(* IEC 61131-3 sources: sis-interlock-demo/pytests/golden/mini/src/GVLs/Generated, 3 files *)

(* ---- GVL_Sis.gvl.st ---- *)
// AUTO-GENERATED by cemgen 1.0.0 — не редактировать: правьте матрицу и запустите
//   python -m cemgen generate <файл матрицы .csv или .xlsx>
// Матрица: TEST-U301-CEM, объект U-301, ревизия 1 от 2026-10-16, SHA-256 сетки 9067fda96ae55e67
// Назначение: экземпляры ПАЗ объекта U-301: источник времени, журнал событий, приложение ПАЗ и
//             команды HMI (ST_SisCmd). Вызов — PRG_Sis.
// Автор:      pytest; код — генератор cemgen
// Версия:     1.0.0
// Документ:   docs/DESIGN.md, раздел «10. Генератор cemgen»; docs/cause_effect_matrix.md
// ВНИМАНИЕ:   код демонстрационный и не предназначен для систем безопасности. Реальная ПАЗ требует
//             определения SIL, сертифицированных аппаратных и программных средств и валидации по
//             ГОСТ Р МЭК 61511.
{attribute 'qualified_only'}
VAR_GLOBAL
    fbTime : PL.FB_SystemTime;   // монотонное время LTIME (PL.I_TimeSource)
    fbLog  : FB_SisEventLog;     // журнал событий ПАЗ, кольцо GVL_Const.SIS_LOG_SIZE
    fbApp  : FB_SisApp;          // ПАЗ объекта: привязка, голосование, матрица, выходы
    stCmd  : ST_SisCmd;          // команды HMI: сброс, пусковые обходы, байпасы каналов
END_VAR

(* ---- GVL_SisCfg.gvl.st ---- *)
// AUTO-GENERATED by cemgen 1.0.0 — не редактировать: правьте матрицу и запустите
//   python -m cemgen generate <файл матрицы .csv или .xlsx>
// Матрица: TEST-U301-CEM, объект U-301, ревизия 1 от 2026-10-16, SHA-256 сетки 9067fda96ae55e67
// Назначение: конфигурация ПАЗ объекта U-301 из матрицы причин и следствий: номера причин и
//             следствий, шкалы датчиков, матрица CEM_CFG (с CRC) и группы голосования VOTE_CFG.
//             VAR_GLOBAL CONSTANT: с HMI не меняется (решение D-09), правка — только через матрицу
//             и генератор.
// Автор:      pytest; код — генератор cemgen
// Версия:     1.0.0
// Документ:   docs/DESIGN.md, раздел «10. Генератор cemgen»; docs/cause_effect_matrix.md
// ВНИМАНИЕ:   код демонстрационный и не предназначен для систем безопасности. Реальная ПАЗ требует
//             определения SIL, сертифицированных аппаратных и программных средств и валидации по
//             ГОСТ Р МЭК 61511.
{attribute 'qualified_only'}
VAR_GLOBAL CONSTANT
    // Номера причин: индекс i строки матрицы, бит маски i − 1
    CAUSE_TSH301       : UINT := 1;   // Температура высокая
    CAUSE_PSL302       : UINT := 2;   // Давление низкое
    CAUSE_XS303        : UINT := 3;   // Внешний останов
    CAUSE_COUNT        : UINT := 3;   // причин в матрице
    // Номера следствий: индекс j столбца матрицы
    EFFECT_XV301       : UINT := 1;   // Отсечной клапан XV301
    EFFECT_M302        : UINT := 2;   // Насос M302
    EFFECT_COUNT       : UINT := 2;   // следствий в матрице
    // Шкалы датчиков 4–20 мА (инж. ед.) и нормальные токи для демо и тестов
    AI_TT301_LO_EU     : REAL := 0.0;   // TT301: шкала 0…100 °C
    AI_TT301_HI_EU     : REAL := 100.0;
    AI_TT301_NORMAL_MA : REAL := 10.4;   // 40 °C
    // Матрица причин и следствий (DESIGN.md, 4.2, 6.8): маска следствия — «X» в его столбце
    CEM_CFG : ST_CemCfg := (uiCauseCount := 3, uiEffectCount := 2, xStartTripped := FALSE,
        wMatrixCrc := 16#0F15,
        astCause := [
            (xEnable := TRUE, eSource := E_CauseSource.Voting, tDelay := T#1S),                 // 1 TSH301
            (xEnable := TRUE, eSource := E_CauseSource.Voting, tDelay := T#0S,
                xOverrideAllowed := TRUE, tOverrideMax := T#10M, tOverrideClear := T#30S),      // 2 PSL302
            (xEnable := TRUE, eSource := E_CauseSource.External, tDelay := T#500MS),            // 3 XS303
            (xEnable := FALSE),                                                                 // 4 — резерв
            (xEnable := FALSE),                                                                 // 5 — резерв
            (xEnable := FALSE),                                                                 // 6 — резерв
            (xEnable := FALSE),                                                                 // 7 — резерв
            (xEnable := FALSE),                                                                 // 8 — резерв
            (xEnable := FALSE),                                                                 // 9 — резерв
            (xEnable := FALSE),                                                                 // 10 — резерв
            (xEnable := FALSE),                                                                 // 11 — резерв
            (xEnable := FALSE),                                                                 // 12 — резерв
            (xEnable := FALSE),                                                                 // 13 — резерв
            (xEnable := FALSE),                                                                 // 14 — резерв
            (xEnable := FALSE),                                                                 // 15 — резерв
            (xEnable := FALSE)],                                                                // 16 — резерв
        astEffect := [
            (eSafeState := E_SafeState.Closed, wCauseMask := 16#0003),                          // 1 XV301: 1, 2
            (eSafeState := E_SafeState.Stopped, wCauseMask := 16#0006),                         // 2 M302: 2, 3
            (wCauseMask := 0),                                                                  // 3 — резерв
            (wCauseMask := 0),                                                                  // 4 — резерв
            (wCauseMask := 0),                                                                  // 5 — резерв
            (wCauseMask := 0),                                                                  // 6 — резерв
            (wCauseMask := 0),                                                                  // 7 — резерв
            (wCauseMask := 0),                                                                  // 8 — резерв
            (wCauseMask := 0),                                                                  // 9 — резерв
            (wCauseMask := 0),                                                                  // 10 — резерв
            (wCauseMask := 0),                                                                  // 11 — резерв
            (wCauseMask := 0),                                                                  // 12 — резерв
            (wCauseMask := 0),                                                                  // 13 — резерв
            (wCauseMask := 0),                                                                  // 14 — резерв
            (wCauseMask := 0),                                                                  // 15 — резерв
            (wCauseMask := 0)]);                                                                // 16 — резерв
    // Группы голосования по причинам (DESIGN.md, 5); ext — без голосования (eArch := None)
    VOTE_CFG : ARRAY[1..GVL_Const.SIS_CAUSES_MAX] OF ST_VotingCfg := [
        (eArch := E_VoteArch.Vote1oo1, ePolicy := E_DegradePolicy.VoteTrip,
            eInput := E_SisInputKind.Analog, eLimitDir := E_LimitDir.High,
            rTripLimit_eu := 80.0, rHyst_eu := 0.0, rDiscrepancyMax_eu := 0.0,
            tDiscrepancyDelay := T#5S, tBypassMax := T#0S, uiMaxBypass := 0),          // 1 TSH301
        (eArch := E_VoteArch.Vote2oo2, ePolicy := E_DegradePolicy.VoteTrip,
            eInput := E_SisInputKind.Discrete, xDiHealthy := TRUE,
            tBypassMax := T#1H, uiMaxBypass := 1),                                     // 2 PSL302
        (eArch := E_VoteArch.None),                                                    // 3 XS303 — ext, без голосования
        (eArch := E_VoteArch.None),                                                    // 4 — резерв
        (eArch := E_VoteArch.None),                                                    // 5 — резерв
        (eArch := E_VoteArch.None),                                                    // 6 — резерв
        (eArch := E_VoteArch.None),                                                    // 7 — резерв
        (eArch := E_VoteArch.None),                                                    // 8 — резерв
        (eArch := E_VoteArch.None),                                                    // 9 — резерв
        (eArch := E_VoteArch.None),                                                    // 10 — резерв
        (eArch := E_VoteArch.None),                                                    // 11 — резерв
        (eArch := E_VoteArch.None),                                                    // 12 — резерв
        (eArch := E_VoteArch.None),                                                    // 13 — резерв
        (eArch := E_VoteArch.None),                                                    // 14 — резерв
        (eArch := E_VoteArch.None),                                                    // 15 — резерв
        (eArch := E_VoteArch.None)];                                                   // 16 — резерв
END_VAR

(* ---- GVL_SisIo.gvl.st ---- *)
// AUTO-GENERATED by cemgen 1.0.0 — не редактировать: правьте матрицу и запустите
//   python -m cemgen generate <файл матрицы .csv или .xlsx>
// Матрица: TEST-U301-CEM, объект U-301, ревизия 1 от 2026-10-16, SHA-256 сетки 9067fda96ae55e67
// Назначение: образ ввода-вывода ПАЗ объекта U-301. Поля stIo привязываются к каналам модулей
//             ввода-вывода; в демо без ввода-вывода PRG_Main ставит нормальные значения
//             (F_SisIoNormal).
// Автор:      pytest; код — генератор cemgen
// Версия:     1.0.0
// Документ:   docs/DESIGN.md, раздел «10. Генератор cemgen»; docs/cause_effect_matrix.md
// ВНИМАНИЕ:   код демонстрационный и не предназначен для систем безопасности. Реальная ПАЗ требует
//             определения SIL, сертифицированных аппаратных и программных средств и валидации по
//             ГОСТ Р МЭК 61511.
{attribute 'qualified_only'}
VAR_GLOBAL
    stIo : ST_SisIo;   // входы датчиков, ключи, кнопка, выходы-разрешения xQ*
END_VAR
